SUBAPPLICATION AX_TO_BG_PUBLISH_SWITCHPIC_Option (* Reine Anzeige: AX-Zustand auf Hintergrundfarbe (SoftKey+AUX), lokalen State-Publish und ObjectPointer-Statusanzeige, aktiviert per AOption (INIT/QI ueber AOption_X_TO_EVENT, INIT_CNF echt nach ObjPtr.INITO). *)
  (* Standard: 61499-2; Description: Copyright (c) 2026 Meisterschulen am Ostbahnhof This program and the accompanying materials are made available under the terms of the Eclipse Public License 2.0 which is available at https://www.eclipse.org/legal/epl-2.0/ SPDX-License-Identifier: EPL-2.0 *)
  (* Version 1.0, 2026-10-17, Franz Höpfinger, Meisterschulen am Ostbahnhof, initial implementation - Anzeige-Teil von AX_TO_QXA_BG_PUBLISH_SWITCHPIC_OPT als eigener Baustein (Franz: an AOption_OR_2_Anzeige ein reiner Anzeige-Baustein). *)
  PACKAGE MyLib::sys;
  IMPORT isobus::UT::Q::const::IDs::ID_NULL;
  IMPORT isobus::UT::Q::types::s2x1ObjectIDs;
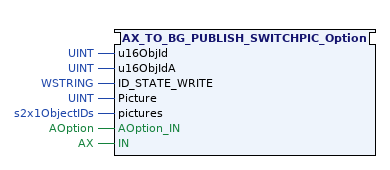
  VAR_INPUT
    u16ObjId : UINT := ID_NULL; (* Object ID Softkey - traegt die Hintergrundfarbe *)
    u16ObjIdA : UINT := ID_NULL; (* Object ID AuxFunction2 (Joystick) - zeigt Hintergrundfarbe am Aux-Handle mit *)
    ID_STATE_WRITE : WSTRING; (* Lokale Publish-Adresse (ACTION=WRITE) fuer den Zustand - wird remote abonniert *)
    Picture : UINT; (* Object ID des ObjectPointer, der den Status-Kaestchen-Inhalt traegt *)
    pictures : isobus::UT::Q::types::s2x1ObjectIDs := (up := (u16ObjId := ID_NULL), down := (u16ObjId := ID_NULL)); (* die beiden Ziel-Object-IDs (up=aus, down=an) *)
  END_VAR
  SOCKETS
    AOption_IN : Option::AOption; (* Aktiviert/deaktiviert die Anzeige *)
    IN : adapter::types::unidirectional::AX; (* Fertiger AX-Zustand fuer Hintergrund, Publish und ObjectPointer *)
  END_SOCKETS
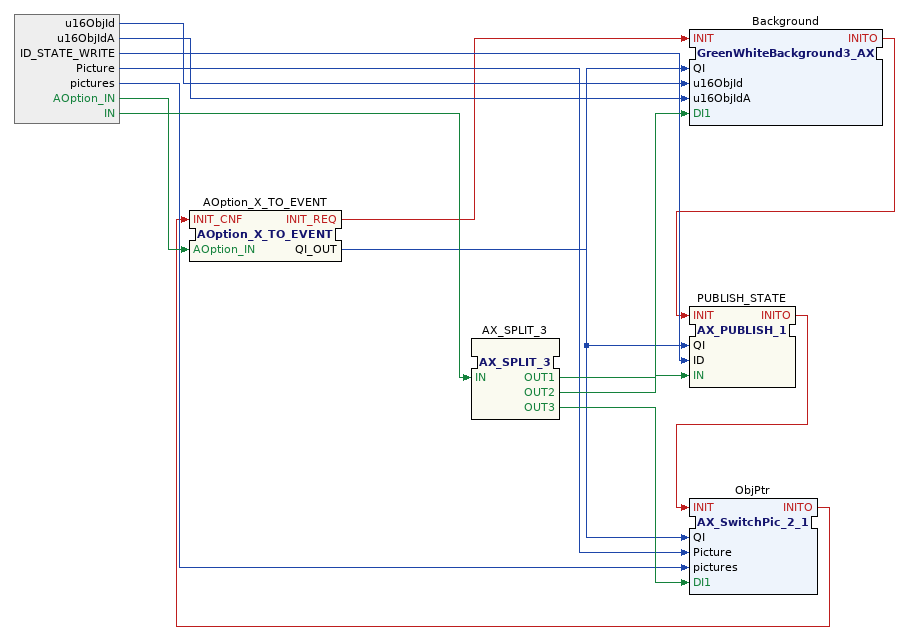
  FBS
    AOption_X_TO_EVENT : Option::conversion::AOption_X_TO_EVENT;
    AX_SPLIT_3 : adapter::events::unidirectional::AX_SPLIT_3; (* Adapter-Fanout ist strikt 1:1 *)
    PUBLISH_STATE : adapter::net::AX_PUBLISH_1;
  END_FBS
  SUBAPPS
    Background : MyLib::sys::GreenWhiteBackground3_AX;
    ObjPtr : MyLib::sys::AX_SwitchPic_2_1;
  END_SUBAPPS
  EVENT_CONNECTIONS
    AOption_X_TO_EVENT.INIT_REQ TO Background.INIT;
    Background.INITO TO PUBLISH_STATE.INIT;
    PUBLISH_STATE.INITO TO ObjPtr.INIT;
    ObjPtr.INITO TO AOption_X_TO_EVENT.INIT_CNF;
  END_CONNECTIONS
  DATA_CONNECTIONS
    AOption_X_TO_EVENT.QI_OUT TO Background.QI;
    AOption_X_TO_EVENT.QI_OUT TO PUBLISH_STATE.QI;
    AOption_X_TO_EVENT.QI_OUT TO ObjPtr.QI;
    u16ObjId TO Background.u16ObjId;
    u16ObjIdA TO Background.u16ObjIdA;
    ID_STATE_WRITE TO PUBLISH_STATE.ID;
    Picture TO ObjPtr.Picture;
    pictures TO ObjPtr.pictures;
  END_CONNECTIONS
  ADAPTER_CONNECTIONS
    AOption_IN TO AOption_X_TO_EVENT.AOption_IN;
    IN TO AX_SPLIT_3.IN;
    AX_SPLIT_3.OUT1 TO Background.DI1;
    AX_SPLIT_3.OUT2 TO PUBLISH_STATE.IN;
    AX_SPLIT_3.OUT3 TO ObjPtr.DI1;
  END_CONNECTIONS
END_SUBAPPLICATION
